TYPE ST_TriggerTellConfiguration :
STRUCT
	bDisableAttention : BOOL;
	commTimeout		  : TIME := T#10S;
END_STRUCT
END_TYPE

(* stored: Version 1.1.0.1, ProductVersion 3.1.4024.12
   DUT ST_TriggerTellConfiguration: Id {4594a0ef-8c32-4939-9647-74d8c847c659} *)
